{region 'Documentation'}
(*!
<summary>Reject a falling edge between consecutive active observations.</summary>
<description>

The first active observation establishes a baseline without deciding a result. Disabling
observation invalidates that baseline, not the held Result. Re-enabling first establishes a new
baseline; Reset clears history.

ObserveFirstCycle FALSE delays the first observation by one enabled call.

</description>
*)
{endregion}
FUNCTION_BLOCK AssertNoFallingEdge EXTENDS AssertionBase
VAR_INPUT
    IN : BOOL; //! Actual value checked or observed by this Assertion.
END_VAR
VAR
    FINPrevious : BOOL;
    FObservationPrevious : BOOL;
    FEvaluationActive : BOOL;
END_VAR

SUPER^();

{region 'Documentation'}
(*!
<summary>Maintain observation history before evaluating the selected edge.</summary>
*)
{endregion}
METHOD PROTECTED Assert
VAR
    PreviousValue : BOOL;
END_VAR
FEvaluationActive := ObservationActive AND FObservationPrevious;
FObservationPrevious := ObservationActive;

IF NOT ObservationActive THEN
    RETURN;
END_IF;

PreviousValue := FINPrevious;
FINPrevious := IN;

IF NOT EvaluationActive THEN
    RETURN;
END_IF;

IF Result = E_Result.Error THEN
    RETURN;
END_IF;

IF Result = E_Result.Failed THEN
    RETURN;
END_IF;

IF NOT IN AND PreviousValue THEN
    Fail(Message := 'Assertion failed: unexpected falling edge detected.');
    RETURN;
END_IF;

Pass();
END_METHOD

{region 'Documentation'}
(*!
<summary>Current/last call can compare two consecutive active observations.</summary>
*)
{endregion}
{attribute 'monitoring' := 'call'}
PROPERTY PUBLIC EvaluationActive : BOOL //! Current/last call can compare two consecutive active observations.
GET // PUBLIC
EvaluationActive := FEvaluationActive;
END_GET
END_PROPERTY

{region 'Documentation'}
(*!
<summary>Clear observation history and the current evaluation gate.</summary>
*)
{endregion}
METHOD PROTECTED ResetAssertion
FINPrevious := FALSE;
FObservationPrevious := FALSE;
FEvaluationActive := FALSE;
END_METHOD

END_FUNCTION_BLOCK

(* stored: Version 1.1.0.1
   POU AssertNoFallingEdge: Id {56a82304-a4d1-464d-951a-1edb78feea88}, SpecialFunc None
   Folder Internal: Id {5365c8a9-4649-4e1d-b5a2-675d8c303ce6}
   Method Assert: Id {64c0943f-9d89-4a3e-ace5-51c0eae664cf}
   Property EvaluationActive: Id {4b27abde-4064-479a-9eda-f349cde88544}
   Get Get: Id {86660a12-81cc-44c4-bd54-1dc0854ad515}
   Method ResetAssertion: Id {8450a173-7994-40ee-aea2-f7edef5229eb} *)
